(* IEC 61131-3 sources: HappyLearnCodesys/content/softmotion/Robotics_Triggers_Advanced, 4 files *)

(* ---- GVL.st ---- *)
{attribute 'qualified_only'}
(*
    檔案用途：
      定義與觸發計時相關的全域常數，包括匯流排週期時間與觸發預測最大時間。
    教學重點：
      - BUS_CYCLE_TIME_IN_US / BUS_CYCLE_TIME_IN_S：提供 TriggerWithTimeShift 參考的基礎時間單位。
      - MAX_TRIGGER_FORECAST_DURATION：根據膠閥與 UV 燈的延遲，自動計算規劃器需要預測的最長時間。
*)
VAR_GLOBAL CONSTANT
    /// 匯流排週期時間（微秒）。
    BUS_CYCLE_TIME_IN_US : DWORD := 4000;
    /// 匯流排週期時間（秒）。
    BUS_CYCLE_TIME_IN_S : LREAL := TO_LREAL(BUS_CYCLE_TIME_IN_US) * 1E-6;
    /// 規劃器需預測的最大觸發時間，取膠閥與 UV 燈延遲的較大值。
    MAX_TRIGGER_FORECAST_DURATION : LREAL := MAX(GlueApplication.GLUE_ON_OFF_DELAY, GlueApplication.UV_LAMP_OFF_DELAY);
END_VAR

(* ---- TriggerWithTimeShift.st ---- *)
(*
    檔案用途：
      封裝 SoftMotion 觸發的「準備、監控與時間位移」邏輯，提供可重複使用的功能塊，
      讓使用者可以指定觸發位置型態與 TimeShift，並取得剩餘觸發時間與觸發狀態。
    教學重點：
      - 比較 STATE_PREPARE_TRIGGER、STATE_MONITOR_TRIGGER、STATE_DECREMENT_REMAINING_TRIGGER_TIME
        等狀態之間的關係，理解如何在每個匯流排週期持續更新 TriggerTime。
      - 注意 TimeShift 為正／負時，TriggerTime 的意義與判斷條件（<= BUS_CYCLE_TIME_IN_S）。
      - 了解 Aborted / Done / Error 等輸出旗標如何反映觸發在實際運行中的各種結束情況。
*)
FUNCTION_BLOCK TriggerWithTimeShift
VAR_IN_OUT
    AxisGroup : AXIS_GROUP_REF_SM3;
END_VAR
VAR_INPUT
    Execute : BOOL;
    PositionType : SMC_TriggerPositionType;
    Position : SMC_TriggerPosition;
    /// The time shift in seconds that the trigger should fire before (positive value)
    /// or after (negative value) the trigger position has been reached.
    /// Please note: Positive time shifts cannot always be met, see the documentation of
    /// ``TriggerTime`` for additional information.
    TimeShift : LREAL;
END_VAR
VAR_OUTPUT
    Busy : BOOL;
    /// The trigger got aborted, i.e. no movement was commanded in the cycle
    /// when the trigger was prepared.
    Aborted : BOOL;
    /// The Trigger is Done in the cycle after the trigger has been reached
    /// or if the movement that the trigger was assigned to got aborted (i.e.
    /// the trigger will never be reached).
    Done : BOOL;
    Error : BOOL;
    ErrorID : SMC_ERROR;
    /// The trigger has been successfully prepared and will be attached to the next
    /// commanded movement.
    TriggerPrepared : BOOL;
    /// The trigger time becomes valid, when the trigger position is part of the known
    /// trajectory.
    TriggerTimeValid : BOOL;
    /// The time in seconds until the trigger position including time shift is reached.
    /// The time is based on the start of the bus task cycle.
    /// Only valid if ``TriggerTimeValid`` is set.
    /// Can be negative, if the time until the trigger position is reached is smaller
    /// than the defined positive time shift. For example, the trigger position is 50 ms
    /// away from the start of the movement, but a positive time shift of 150 ms was
    /// defined. Since the start of the movement does not get delayed, the trigger
    /// will get noticed 100 ms too late.
    TriggerTime : LREAL;
    /// The trigger position including time shift is reached this cycle.
    TriggerReachedThisCycle : BOOL;
END_VAR
VAR
    m_state : INT;

    m_prepareTrigger : SMC_GroupPrepareTrigger;
    m_readTrigger : SMC_GroupReadTrigger;

    m_oldExecute : BOOL;
END_VAR
VAR_TEMP
    triggerTimeWithoutTimeShift : LREAL;
END_VAR
VAR CONSTANT
    STATE_IDLE : INT := 0;
    STATE_PREPARE_TRIGGER : INT := 10;
    STATE_MONITOR_TRIGGER : INT := 20;
    STATE_DECREMENT_REMAINING_TRIGGER_TIME : INT := 30;
    STATE_TRIGGER_FIRED : INT := 100;
    STATE_DONE : INT := 500;
    STATE_ABORTED : INT := 600;
    STATE_ERROR : INT := 1000;
END_VAR

IF Execute AND NOT m_oldExecute THEN
    m_prepareTrigger(
        AxisGroup:= AxisGroup,
        Execute:= FALSE);
    m_readTrigger(
        AxisGroup:= AxisGroup,
        Enable:= FALSE);

    m_state := STATE_PREPARE_TRIGGER;
ELSIF NOT Execute AND (Done OR Error OR Aborted) THEN
    m_state := STATE_IDLE;
    ErrorID := SMC_NO_ERROR;
END_IF

CASE m_state OF
STATE_PREPARE_TRIGGER:
    m_prepareTrigger(
        AxisGroup:= AxisGroup,
        Execute:= TRUE,
        PositionType:= PositionType,
        Position:= Position);

    IF m_prepareTrigger.Done THEN
        m_state := STATE_MONITOR_TRIGGER;
    ELSIF m_prepareTrigger.Error THEN
        m_state := STATE_ERROR;
        ErrorID := m_prepareTrigger.ErrorID;
    ELSIF m_prepareTrigger.CommandAborted THEN
        m_state := STATE_ABORTED;
    END_IF

STATE_MONITOR_TRIGGER:
    m_readTrigger(
        AxisGroup:= AxisGroup,
        Enable:= TRUE,
        TriggerId:= m_prepareTrigger.TriggerId);

    IF m_readTrigger.TriggerInfo.status = SMC_TRIGGER_STATUS.Active THEN
        triggerTimeWithoutTimeShift := m_readTrigger.TriggerInfo.triggerTime;
        TriggerTime := triggerTimeWithoutTimeShift - TimeShift;

        IF TriggerTime <= GVL.BUS_CYCLE_TIME_IN_S THEN
            m_state := STATE_TRIGGER_FIRED;
        ELSIF triggerTimeWithoutTimeShift <= GVL.BUS_CYCLE_TIME_IN_S THEN
            m_state := STATE_DECREMENT_REMAINING_TRIGGER_TIME;
        END_IF
    ELSIF m_readTrigger.TriggerInfo.status = SMC_TRIGGER_STATUS.Error THEN
        m_state := STATE_ERROR;
        ErrorID := m_readTrigger.TriggerInfo.errorId;
    ELSIF m_readTrigger.TriggerInfo.status <> SMC_TRIGGER_STATUS.Enabled THEN
        /// The movement that the trigger was assigned to got aborted.
        /// The trigger will never be reached. Switch to Done.
        m_state := STATE_DONE;
    END_IF

STATE_DECREMENT_REMAINING_TRIGGER_TIME:
    TriggerTime := TriggerTime - GVL.BUS_CYCLE_TIME_IN_S;
    IF TriggerTime <= GVL.BUS_CYCLE_TIME_IN_S THEN
        m_state := STATE_TRIGGER_FIRED;
    END_IF

STATE_TRIGGER_FIRED:
    m_state := STATE_DONE;
    TriggerTime := 0;
END_CASE

Busy := m_state > STATE_IDLE AND m_state < STATE_DONE;
TriggerPrepared := m_prepareTrigger.Prepared AND m_state > STATE_IDLE;
TriggerTimeValid :=
    m_state = STATE_MONITOR_TRIGGER AND m_readTrigger.TriggerInfo.status = SMC_TRIGGER_STATUS.Active
    OR m_state = STATE_DECREMENT_REMAINING_TRIGGER_TIME
    OR m_state = STATE_TRIGGER_FIRED;
TriggerReachedThisCycle := m_state = STATE_TRIGGER_FIRED;
Aborted := m_state = STATE_ABORTED;
Done := m_state = STATE_DONE;
Error := m_state = STATE_ERROR;

m_oldExecute := Execute;

(* ---- GlueApplication.st ---- *)
(*
    檔案用途：
      模擬一個「點膠＋UV 固化」的應用範例，控制二軸平面運動，同時配合多個觸發點
      來開關膠閥、UV 燈與膠料補充訊號。
    教學重點：
      - 了解如何將一連串線性運動切成多段（GLUE_POSITIONS），並在特定段落上掛載 TriggerWithTimeShift。
      - 觀察不同 PositionType（MvtRelative、MvtDistance、PlaneIntersection）與 TimeShift 正負值的用法。
      - 練習從狀態機 m_state 的角度閱讀「初始化 → 上電 → 多段運動＋觸發 → 監控觸發 → 結束」的流程。
*)
PROGRAM GlueApplication
VAR_OUTPUT
    EnableGlue : BOOL;
    EnableUVLamp : BOOL;
    RefillGlueStorage : BOOL;
END_VAR
VAR
    m_state : INT;
    m_groupPower : SMC_GroupPower;
    m_groupEnable : MC_GroupEnable;

    m_moveLinearAbsolutes : ARRAY[0..MOVEMENT_COUNT - 1] OF MC_MoveLinearAbsolute;

    m_enableGlueTrigger : TriggerWithTimeShift;
    m_disableGlueTrigger : TriggerWithTimeShift;
    m_refillGlueStorageTrigger : TriggerWithTimeShift;
    m_enableUVLampTrigger : TriggerWithTimeShift;
    m_disableUVLampTrigger : TriggerWithTimeShift;
END_VAR
VAR CONSTANT
    MOVEMENT_COUNT : UINT := 5;

    /// The delay in seconds between starting the glue tool and
    /// the first contact with the surface or the delay between
    /// stopping the glue tool and the stop of contact with the
    /// surface.
    GLUE_ON_OFF_DELAY : LREAL := 0.05;
    /// The delay in seconds when the UV-lamp should turn off
    /// after applying glue to the surface. Has to be negative
    /// for the trigger to fire after the position has been
    /// passed.
    UV_LAMP_OFF_DELAY : LREAL := -1.5;

    GLUE_POSITIONS : ARRAY[0..MOVEMENT_COUNT - 1] OF SMC_POS_REF :=
        [
            (c:= (X:= 10)),
            (c:= (X:= 10, Y:= 2)),
            (c:= (X:= 0, Y:= 2)),
            (c:= (X:= 0, Y:= 4)),
            (c:= (X:= 10, Y:= 4))
        ];

    STATE_INIT : INT := 0;
    STATE_POWER_AND_ENABLE : INT := 10;
    STATE_COMMAND_FIRST_MOVEMENT_WITH_TRIGGERS : INT := 20;
    STATE_COMMAND_SECOND_MOVEMENT : INT := 30;
    STATE_COMMAND_THIRD_MOVEMENT_WITH_TRIGGERS : INT := 40;
    STATE_COMMAND_FOURTH_MOVEMENT : INT := 50;
    STATE_COMMAND_FIFTH_MOVEMENT_WITH_TRIGGERS : INT := 60;
    STATE_MONITOR_MOVEMENTS_AND_TRIGGERS : INT := 70;
    STATE_DONE : INT := 500;
END_VAR

CASE m_state OF
STATE_INIT:
    IF Planning_PRG.initDone THEN
        InitializeMovementPOUs();
        m_state := STATE_POWER_AND_ENABLE;
    END_IF

STATE_POWER_AND_ENABLE:
    m_groupPower.Enable := TRUE;
    m_groupPower.bDriveStart := TRUE;
    m_groupPower.bRegulatorOn := TRUE;

    m_groupEnable.Execute := m_groupPower.Status;

    IF m_groupPower.Status AND m_groupEnable.Done THEN
        m_state := STATE_COMMAND_FIRST_MOVEMENT_WITH_TRIGGERS;
    END_IF

STATE_COMMAND_FIRST_MOVEMENT_WITH_TRIGGERS:
    m_enableGlueTrigger.Position.MvtPosition := 0.5;
    m_enableGlueTrigger.PositionType := SMC_TriggerPositionType.MvtRelative;
    m_enableGlueTrigger.TimeShift := GLUE_ON_OFF_DELAY;
    m_enableGlueTrigger(AxisGroup:= AxisGroup, Execute:= TRUE);

    m_enableUVLampTrigger.Position.MvtPosition := 0.5;
    m_enableUVLampTrigger.PositionType := SMC_TriggerPositionType.MvtRelative;
    m_enableUVLampTrigger(AxisGroup:= AxisGroup, Execute:= TRUE);

    m_moveLinearAbsolutes[0](
        AxisGroup:= AxisGroup,
        Execute:= m_enableGlueTrigger.TriggerPrepared AND m_enableUVLampTrigger.TriggerPrepared);

    IF m_moveLinearAbsolutes[0].CommandAccepted THEN
        m_state := STATE_COMMAND_SECOND_MOVEMENT;
    END_IF

STATE_COMMAND_SECOND_MOVEMENT:
    m_moveLinearAbsolutes[1](AxisGroup:= AxisGroup, Execute:= TRUE);

    IF m_moveLinearAbsolutes[1].CommandAccepted THEN
        m_state := STATE_COMMAND_THIRD_MOVEMENT_WITH_TRIGGERS;
    END_IF

STATE_COMMAND_THIRD_MOVEMENT_WITH_TRIGGERS:
    m_refillGlueStorageTrigger.Position.MvtPosition := 5;
    m_refillGlueStorageTrigger.PositionType := SMC_TriggerPositionType.MvtDistance;
    m_refillGlueStorageTrigger(AxisGroup:= AxisGroup, Execute:= TRUE);

    m_moveLinearAbsolutes[2](
        AxisGroup:= AxisGroup,
        Execute:= m_refillGlueStorageTrigger.TriggerPrepared);

    IF m_moveLinearAbsolutes[2].CommandAccepted THEN
        m_state := STATE_COMMAND_FOURTH_MOVEMENT;
    END_IF

STATE_COMMAND_FOURTH_MOVEMENT:
    m_moveLinearAbsolutes[3](AxisGroup:= AxisGroup, Execute:= TRUE);

    IF m_moveLinearAbsolutes[3].CommandAccepted THEN
        m_state := STATE_COMMAND_FIFTH_MOVEMENT_WITH_TRIGGERS;
    END_IF

STATE_COMMAND_FIFTH_MOVEMENT_WITH_TRIGGERS:
    m_disableGlueTrigger.Position.Plane.CoordSystem := SMC_COORD_SYSTEM.MCS;
    m_disableGlueTrigger.Position.Plane.Distance := 5;
    m_disableGlueTrigger.Position.Plane.NormalVector.dX := 1;
    m_disableGlueTrigger.PositionType := SMC_TriggerPositionType.PlaneIntersection;
    m_disableGlueTrigger.TimeShift := GLUE_ON_OFF_DELAY;
    m_disableGlueTrigger(AxisGroup:= AxisGroup, Execute:= TRUE);

    m_disableUVLampTrigger.Position := m_disableGlueTrigger.Position;
    m_disableUVLampTrigger.PositionType := SMC_TriggerPositionType.PlaneIntersection;
    m_disableUVLampTrigger.TimeShift := UV_LAMP_OFF_DELAY;
    m_disableUVLampTrigger(AxisGroup:= AxisGroup, Execute:= TRUE);

    m_moveLinearAbsolutes[4](
        AxisGroup:= AxisGroup,
        Execute:= m_disableGlueTrigger.TriggerPrepared AND m_disableUVLampTrigger.TriggerPrepared);

    IF m_moveLinearAbsolutes[4].CommandAccepted THEN
        m_state := STATE_MONITOR_MOVEMENTS_AND_TRIGGERS;
    END_IF

STATE_MONITOR_MOVEMENTS_AND_TRIGGERS:
    CallTriggers();
    EvaluateTriggers();

    IF m_moveLinearAbsolutes[MOVEMENT_COUNT - 1].Done
       AND NOT EnableGlue
       AND NOT EnableUVLamp
       AND NOT RefillGlueStorage
    THEN
        m_state := STATE_DONE;
    END_IF
END_CASE

m_groupPower(AxisGroup:= AxisGroup);
m_groupEnable(AxisGroup:= AxisGroup);
CallMovements();

(* ---- Planning_PRG.st ---- *)
(*
    檔案用途：
      與基礎 Triggers 範例類似，在規劃任務中呼叫 SMC_TuneCPKernel，
      但這裡的預測時間 fPlanningForecastDuration 根據 GVL.MAX_TRIGGER_FORECAST_DURATION 動態決定，
      以涵蓋膠閥與 UV 燈兩種不同延遲的最大值。
    教學重點：
      - 從觸發應用的角度理解「規劃器預測時間」與「周邊設備延遲」之間的關係。
      - 認識如何透過 GVL 將機台整體時序需求集中配置，再由 Planning_PRG 套用到規劃核心。
*)
PROGRAM Planning_PRG
VAR_OUTPUT
    initDone : BOOL;
END_VAR
VAR
    tuneCPKernel : SMC_TuneCPKernel;
END_VAR

tuneCPKernel(
    AxisGroup:= AxisGroup,
    Execute:= TRUE,
    fPlanningForecastDuration:= GVL.MAX_TRIGGER_FORECAST_DURATION);

initDone := tuneCPKernel.Done;
